// TIA Portal V20 export
// export: Created 2026-10-12T16:46:22.8826847Z, ExportSetting WithDefaults, DisplayName Totally Integrated Automation Portal, DisplayVersion V20 Update 6, DisplayName TIA Portal Openness, DisplayVersion V20 Update 6, DisplayName TIA Portal Version Control Interface, DisplayVersion V20 Update 6, DisplayName SINAMICS Startdrive Advanced, DisplayVersion V20 SP1 Update 2, DisplayName SINAMICS Startdrive G110M, G120, G120C, G120D, G120P, G115D, DisplayVersion V20 SP1 Update 2, DisplayName SINAMICS Startdrive G130, G150, S120, S150, SINAMICS MV, G220, S200, S210, DisplayVersion V20 SP1 Update 2, DisplayName STEP 7 Professional, DisplayVersion V20 Update 6, DisplayName STEP 7 Safety, DisplayVersion V20 Update 2, DisplayName WinCC Basic/Comfort/Advanced, DisplayVersion V20 Update 6, DisplayName WinCC Professional, DisplayVersion V20 Update 6, DisplayName WinCC Unified, DisplayVersion V20 Update 6
TYPE "UDT_BadStatus"
// stored: IsFailsafeCompliant false
   STRUCT
      Belegt : Bool;   // Bad ist belegt
      Auftragsindex : Int;   // Welcher Auftrag belegt dieses Bad
      SchrittIndex : Int;   // Welcher Schritt im Auftrag
      Istzeit : Time;   // Bereits verstrichene Zeit
      Restzeit : Time;   // Verbleibende Verweilzeit
      Zeit_Abgelaufen : Bool;   // Verweilzeit erreicht
      Krit_Zeit_Abgelaufen : Bool;   // Kritische Zeit überschritten
      Ampel_Status : Int;   // 0=Aus, 1=GrünBlink(warte auf WT-Einsetzen), 2=Grün(belegt,OK), 3=GelbBlink(Vorwarnung), 4=RotBlink(Zeit über), 5=RotBlink+Akustik(krit.Zeit), 6=Rot(nicht betriebsbereit)
      Hupe : Bool;   // Akustischer Alarm aktiv
      WT_Eingesetzt : Bool;   // Bediener hat WT eingesetzt
      WT_Entnommen : Bool;   // Bediener hat WT entnommen
      Betriebsbereit : Bool;   // Bad ist betriebsbereit (Temp, Pumpe, Niveau OK)
   END_STRUCT;
END_TYPE
